Yaskawa INFORM job: 2209_2.JBI

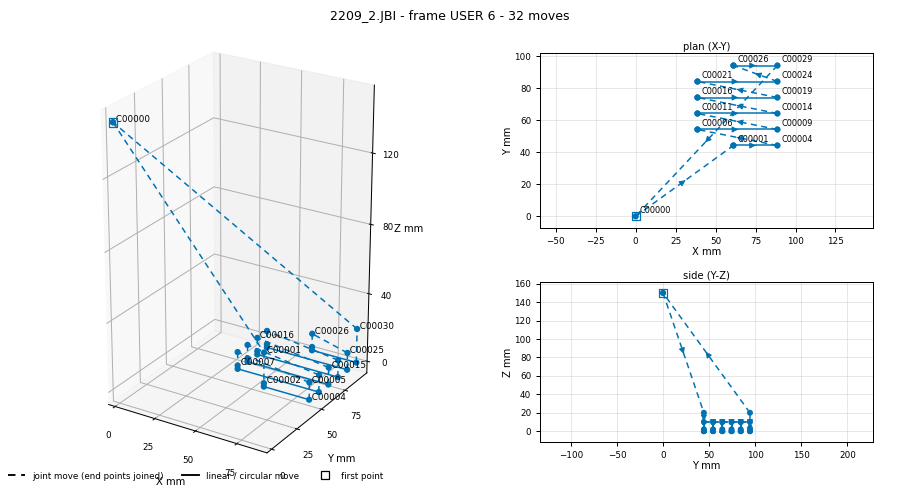
[picture p0: tool path of 2209_2.JBI in frame USER 6, 32 of 32 moves have a stored position in this frame; points joined in program order, loops and branches not executed]
/JOB
//NAME 2209_2
//POS
///NPOS 32,0,0,0,0,0
///USER 6
///TOOL 1
///POSTYPE USER
///RECTAN
///RCONF 1,0,0,0,0,0,0,0,0,0,0,0,0,0,0,0,0,0,0,0,0,0,0,0
C00000=0.000,0.000,150.000,0.0000,0.0000,-50.0000
C00001=61.167,44.319,20.000,0.0000,0.0000,-50.0000
C00002=61.167,44.319,2.000,0.0000,0.0000,-50.0000
C00003=61.167,44.319,0.000,0.0000,0.0000,-50.0000
C00004=88.688,44.319,0.000,0.0000,0.0000,-50.0000
C00005=88.688,44.319,10.000,0.0000,0.0000,-50.0000
C00006=38.688,54.319,10.000,0.0000,0.0000,-50.0000
C00007=38.688,54.319,2.000,0.0000,0.0000,-50.0000
C00008=38.688,54.319,0.000,0.0000,0.0000,-50.0000
C00009=88.688,54.319,0.000,0.0000,0.0000,-50.0000
C00010=88.688,54.319,10.000,0.0000,0.0000,-50.0000
C00011=38.688,64.319,10.000,0.0000,0.0000,-50.0000
C00012=38.688,64.319,2.000,0.0000,0.0000,-50.0000
C00013=38.688,64.319,0.000,0.0000,0.0000,-50.0000
C00014=88.688,64.319,0.000,0.0000,0.0000,-50.0000
C00015=88.688,64.319,10.000,0.0000,0.0000,-50.0000
C00016=38.688,74.319,10.000,0.0000,0.0000,-50.0000
C00017=38.688,74.319,2.000,0.0000,0.0000,-50.0000
C00018=38.688,74.319,0.000,0.0000,0.0000,-50.0000
C00019=88.688,74.319,0.000,0.0000,0.0000,-50.0000
C00020=88.688,74.319,10.000,0.0000,0.0000,-50.0000
C00021=38.688,84.319,10.000,0.0000,0.0000,-50.0000
C00022=38.688,84.319,2.000,0.0000,0.0000,-50.0000
C00023=38.688,84.319,0.000,0.0000,0.0000,-50.0000
C00024=88.688,84.319,0.000,0.0000,0.0000,-50.0000
C00025=88.688,84.319,10.000,0.0000,0.0000,-50.0000
C00026=61.206,94.319,10.000,0.0000,0.0000,-50.0000
C00027=61.206,94.319,2.000,0.0000,0.0000,-50.0000
C00028=61.206,94.319,0.000,0.0000,0.0000,-50.0000
C00029=88.688,94.319,0.000,0.0000,0.0000,-50.0000
C00030=88.688,94.319,20.000,0.0000,0.0000,-50.0000
C00031=0.000,0.000,150.000,0.0000,0.0000,-50.0000
//INST
///DATE 2026/09/22 15:35
///ATTR SC,RW,RJ
////FRAME USER 6
///GROUP1 RB1
NOP
MOVJ C00000 VJ=0.78
MOVJ C00001 VJ=0.78
MOVJ C00002 VJ=0.78
MOVL C00003 V=10.0
MACRO1 MJ#(0) ARGF207
ARCON
MOVL C00004 V=10.0
ARCOF
MOVJ C00005 VJ=0.78
MOVJ C00006 VJ=0.78
MOVJ C00007 VJ=0.78
MOVL C00008 V=10.0
MACRO1 MJ#(0) ARGF207
ARCON
MOVL C00009 V=10.0
ARCOF
MOVJ C00010 VJ=0.78
MOVJ C00011 VJ=0.78
MOVJ C00012 VJ=0.78
MOVL C00013 V=10.0
MACRO1 MJ#(0) ARGF207
ARCON
MOVL C00014 V=10.0
ARCOF
MOVJ C00015 VJ=0.78
MOVJ C00016 VJ=0.78
MOVJ C00017 VJ=0.78
MOVL C00018 V=10.0
MACRO1 MJ#(0) ARGF207
ARCON
MOVL C00019 V=10.0
ARCOF
MOVJ C00020 VJ=0.78
MOVJ C00021 VJ=0.78
MOVJ C00022 VJ=0.78
MOVL C00023 V=10.0
MACRO1 MJ#(0) ARGF207
ARCON
MOVL C00024 V=10.0
ARCOF
MOVJ C00025 VJ=0.78
MOVJ C00026 VJ=0.78
MOVJ C00027 VJ=0.78
MOVL C00028 V=10.0
MACRO1 MJ#(0) ARGF207
ARCON
MOVL C00029 V=10.0
ARCOF
MOVJ C00030 VJ=0.78
MOVJ C00031 VJ=0.78
END
